Fanuc KAREL source: KT00386.KL

PROGRAM KT00386
%NOLOCKGROUP
VAR
  P1: POSITION
  P2: JOINTPOS
  OUT: BOOLEAN
BEGIN
  OUT = P1 <= P2
END KT00386
